FUNCTION_BLOCK FB_DomeErrorState EXTENDS  FB_DomeState
VAR
END_VAR


METHOD CloseCommand : BOOL
// #202: a close is accepted in every state, it is the way to shut the roof
// the error is cleared like a reset does it: the shutter command must not wait for a dome_reset
ResetCommand();
pDome^.SetState(pDome^.fbDomeCloseingState);
END_METHOD


METHOD ResetCommand : BOOL
VAR
	fbClearTx			: ClearComBuffer;
	fbClearRx			: ClearComBuffer;
END_VAR
fbClearTx(Buffer:=TxBuffer);
fbClearRx(Buffer:=TxBuffer);

pDome^._Error := FALSE;
pDome^.SetState(pDome^.fbDomeIdleState);
END_METHOD


PROPERTY StateID : STRING
GET
StateID := 'Error State';
END_GET
END_PROPERTY

END_FUNCTION_BLOCK

(* stored: Version 1.1.0.1, ProductVersion 3.1.4024.15
   POU FB_DomeErrorState: Id {1c3fd2da-883e-4dfd-9e70-6396fe4dc63e}, SpecialFunc None
   Method CloseCommand: Id {2211e3ad-15ee-4774-946f-138090512f81}
   Method ResetCommand: Id {f76344eb-46e9-441e-956f-e4feed1005b3}
   Property StateID: Id {f76a3fa6-76fb-4d56-aec9-546023ad0ca7}
   Get Get: Id {131512d7-c6aa-4508-ab7e-7f04233ba0cb} *)
